Staubli VAL3: Appli_FG_1.pjx

--- Appli_FG_1.pjx ---
Parameters version=s8.15.1Cs9_BS3177 stackSize=200000 millimeterUnit=true
Program file=BP_Validation.pgx
Program file=exercice2.pgx
Program file=exercice3.pgx
Program file=exercice4.pgx
Program file=exercice5.pgx
Program file=exercice6.pgx
Program file=fermerPince.pgx
Program file=IHM.pgx
Program file=Init_Repere.pgx
Program file=ouvrirPince.pgx
Program file=start.pgx
Program file=stop.pgx
Data file=Appli_FG_1.dtx

--- Appli_FG_1.dtx ---
jointRx jDepart = {j3=90, j5=90, j6=90}
mdesc mLent = {vel=10, blend=off}
mdesc mNomSpeed
mdesc mRapide = {vel=25, blend=off}
pointRx Prise5[5]
  [0] = {x=431.0804335, y=26.782897, z=-154.648647, rx=179.571045, ry=-2.0767627, rz=-88.582368, fatherId=world[0]}
  [1] = {x=447.943291, y=66.6588, z=-153.242684, rx=179.468283, ry=-1.214183, rz=-87.886126, fatherId=world[0]}
  [2] = {x=443.413957, y=103.41072, z=-155.933715, rx=179.299339, ry=-1.959881, rz=-87.727854, fatherId=world[0]}
  [3] = {x=442.540779, y=142.243832, z=-156.250835, rx=179.370693, ry=-1.0627126, rz=-86.483272, fatherId=world[0]}
  [4] = {x=448.0116706, y=178.916845, z=-155.959372, rx=178.810182, ry=0.0453744, rz=-89.949172, fatherId=world[0]}
pointRx pDepose = {x=103.42949, y=-354.0596717, z=-68.418859, rx=-176.797277, ry=-1.191891, rz=1.0467852, fatherId=world[0]}
tool tPince = {z=120, fatherId=flange[0], ioLink=ValveIO\valve1}
bool bStart
string nCouleur_Autorisation
frame fcaisse = {fatherId=world[0]}
pointRx plA = {x=5, y=100, z=23, rx=-180, fatherId=fcaisse[0]}
pointRx pRcaisse[3]
  [0] = {x=519.439885783333, y=-120.149697377671, z=-165.099001775512, rx=-179.999991526125, ry=6.52832163301057E-07, rz=3.27642281379904E-06, fatherId=world[0]}
  [1] = {x=519.439876404586, y=139.850292212372, z=-165.098973789677, rx=-179.999991372113, ry=-1.03012204155165E-07, rz=4.01298181690715E-06, fatherId=world[0]}
  [2] = {x=319.439927962114, y=-120.149711900373, z=-165.098985799063, rx=-179.999992133117, ry=1.76060323841222E-06, rz=3.02670493493255E-06, fatherId=world[0]}
bool bInit_repere

--- start.pgx ---
program start()
begin
  resetMotion(jDepart)
  bInit_repere = false
  taskCreate "IHM",10,IHM()
  call exercice6()
end

--- BP_Validation.pgx ---
program BP_Validation()
begin
  bStart[0] = true
end

--- exercice2.pgx ---
program exercice2()
begin
  movej(jDepart,tPince,mRapide)
  call ouvrirPince()
  movej(appro(Prise5[0],{0,0,-50,0,0,0}),tPince,mRapide)
  movel(Prise5[0],tPince,mLent)
  call fermerPince()
  movel(appro(Prise5[0],{0,0,-50,0,0,0}),tPince,mRapide)

  movej(jDepart,tPince,mRapide)
  movej(appro(pDepose[0],{0,0,-50,0,0,0}),tPince,mRapide)
  movel(pDepose[0],tPince,mLent)
  call ouvrirPince()
  movel(appro(pDepose,{0,0,-50,0,0,0}),tPince,mRapide)

  movej(jDepart,tPince,mLent)

  waitEndMove()
end

--- exercice3.pgx ---
program exercice3()
  local num l_n1
begin
  movej(jDepart,tPince,mRapide)
  call ouvrirPince()

  for l_n1 = 0 to 4
    movej(appro(Prise5[l_n1],{0,0,-50,0,0,0}),tPince,mRapide)
    movel(Prise5[l_n1],tPince,mLent)
    call fermerPince()
    movel(appro(Prise5[l_n1],{0,0,-50,0,0,0}),tPince,mRapide)

    movej(jDepart,tPince,mRapide)
    movej(appro(pDepose[0],{0,0,-50,0,0,0}),tPince,mRapide)
    movel(pDepose[0],tPince,mLent)
    call ouvrirPince()
    movel(appro(pDepose,{0,0,-50,0,0,0}),tPince,mRapide)


    movej(jDepart,tPince,mLent)
    waitEndMove()
    delay(3)
  endFor

end

--- exercice4.pgx ---
program exercice4()
  local num l_nNbKapla
  local pointRx dest
  local trsf Pas
  local trsf Decal
begin
  Pas.x = (((Prise5[4].trsf.x)-(Prise5[0].trsf.x))/4)
  Pas.y = (((Prise5[4].trsf.y)-(Prise5[0].trsf.y))/4)
  Pas.z = (((Prise5[4].trsf.z)-(Prise5[0].trsf.z))/4)

  for l_nNbKapla = 0 to 4

    Decal.x = l_nNbKapla * Pas.x
    Decal.y = l_nNbKapla * Pas.y
    Decal.z = l_nNbKapla * Pas.z

    dest = compose(Prise5[0],world,Decal)

    movej(appro(dest,{0,0,-50,0,0,0}),tPince,mRapide)
    movel(dest,tPince,mLent)
    call fermerPince()
    movel(appro(dest,{0,0,-50,0,0,0}),tPince,mRapide)

    movej(jDepart,tPince,mRapide)
    movej(appro(pDepose[0],{0,0,-50,0,0,0}),tPince,mRapide)
    movel(pDepose[0],tPince,mLent)
    call ouvrirPince()
    movel(appro(pDepose,{0,0,-50,0,0,0}),tPince,mRapide)
    movej(jDepart,tPince,mLent)
    waitEndMove()
    delay(3)
    endFor

end

--- exercice5.pgx ---
program exercice5()
  local num l_nNbKapla
  local pointRx dest
  local trsf Pas
  local trsf Decal
begin
  Pas.x = (((Prise5[4].trsf.x)-(Prise5[0].trsf.x))/4)
  Pas.y = (((Prise5[4].trsf.y)-(Prise5[0].trsf.y))/4)
  Pas.z = (((Prise5[4].trsf.z)-(Prise5[0].trsf.z))/4)

  for l_nNbKapla = 0 to 4

    Decal.x = l_nNbKapla * Pas.x
    Decal.y = l_nNbKapla * Pas.y
    Decal.z = l_nNbKapla * Pas.z

    dest = compose(Prise5[0],world,Decal)

    bStart = false
    nCouleur_Autorisation = "#80EA34"
    movej(appro(dest,{0,0,-50,0,0,0}),tPince,mRapide)
    movel(dest,tPince,mLent)
    call fermerPince()
    movel(appro(dest,{0,0,-50,0,0,0}),tPince,mRapide)
    movej(jDepart,tPince,mRapide)


    wait(bStart == true)


    nCouleur_Autorisation = "#EA3734"
    movej(appro(pDepose[0],{0,0,-50,0,0,0}),tPince,mRapide)
    movel(pDepose[0],tPince,mLent)
    call ouvrirPince()
    movel(appro(pDepose[0],{0,0,-50,0,0,0}),tPince,mRapide)
    movej(jDepart,tPince,mLent)
    waitEndMove()


  endFor
end

--- exercice6.pgx ---
program exercice6()
  local num l_nNbKapla
  local pointRx dest
  local trsf Pas
  local trsf Decal
begin

  wait(bInit_repere == true)
  for l_nNbKapla = 0 to 4

    Decal.x = l_nNbKapla * 40

    dest = compose(plA,fcaisse,Decal)

    bStart = false
    nCouleur_Autorisation = "#80EA34"
    movej(appro(dest,{0,0,-50,0,0,0}),tPince,mRapide)
    movel(dest,tPince,mLent)
    call fermerPince()
    movel(appro(dest,{0,0,-50,0,0,0}),tPince,mRapide)
    movej(jDepart,tPince,mRapide)

    wait(bStart == true)
    nCouleur_Autorisation = "#EA3734"
    movej(appro(pDepose[0],{0,0,-50,0,0,0}),tPince,mRapide)
    movel(pDepose[0],tPince,mLent)
    call ouvrirPince()
    movel(appro(pDepose[0],{0,0,-50,0,0,0}),tPince,mRapide)
    movej(jDepart,tPince,mLent)
    waitEndMove()


  endFor
end

--- fermerPince.pgx ---
program fermerPince()
begin
  open(tPince)
end

--- IHM.pgx ---
program IHM()
begin
  userPage("IHM")
  while true
    delay(0.5)
  endWhile
end

--- Init_Repere.pgx ---
program Init_Repere()
begin
  bInit_repere =true
  setFrame(pRcaisse[0], pRcaisse[1], pRcaisse[2],fcaisse)
end

--- ouvrirPince.pgx ---
program ouvrirPince()
begin
  close(tPince)
end

--- stop.pgx ---
program stop()
begin
end
